(* IEC 61131-3 sources: PLC-Static-Analysis/modules/plc-rules/src/test/resources/PLCA-L025, 2 files *)

(* ---- compliant.st ---- *)
PROGRAM P_L025ok
VAR
    n : INT;
    m : INT;
    r : REAL;
    b : BOOL;
    c : BOOL;
    q : BOOL;
END_VAR
IF b THEN
    q := FALSE;
END_IF
q := b = c;
q := n = 1;
END_PROGRAM

(* ---- noncompliant.st ---- *)
PROGRAM P_L025
VAR
    n : INT;
    m : INT;
    r : REAL;
    b : BOOL;
    c : BOOL;
    q : BOOL;
END_VAR
IF b = TRUE THEN // PLCA-L025
    q := FALSE;
END_IF
q := c <> FALSE; // PLCA-L025
q := FALSE = (n > 3); // PLCA-L025
END_PROGRAM
